FUNCTION_BLOCK FB_ScalingOffset_1
(*

The function block used to scaling input signal.

Constructor: 		Patryk Panylo
Company:		E. Riexinger GmbH
Date:			04.08.2015
Version:			1.00

Date:			Revision:		Who:				Comment
dd.mm.yyyy		x.xx			Initials			comment

*)
VAR_INPUT
	(* Input variables / Eingang Variablen *)
	bEnable							:BOOL;						(* Function block enable *)
	lrInput							:LREAL;						(* Input scaling proces value *)
	lrXLowLimit						:LREAL;						(* Upper limit of X range *)
	lrXUpperLimit						:LREAL; 						(*Upper limit of X range  *)
	lrYLowLimit						:LREAL; 						(* Low limit of Y range  *)
	lrYUpperLimit						:LREAL; 						(* Upper limit of Y range  *)
	usiPrecision						:USINT := 2; 					(* The number of digits after the decimal point depends on the requested precision *)
	lrOffset							:LREAL;						(* Offset of output *)
END_VAR
VAR_OUTPUT
	(* Output variables / Ausgang Variablen *)
	lrOutputRV						:LREAL;						(* Raw Value *)
	lrOutputPV						:LREAL;						(* Judgment Value  *)
END_VAR
VAR
	(* Instances / Instanzen *)
	fbScaling						:FB_Scaling;

	(* Enumerator  *)

	(* General flags / Allgemeine Variablen *)

END_VAR
VAR CONSTANT

END_VAR

IF NOT bEnable THEN
	fbScaling(
		bEnable := FALSE,
	);

	lrOutputRV := 0.0;					(* Raw Value *)
	lrOutputPV := 0.0;					(* Judgment Value *)
	RETURN;
END_IF

(* Scaling *)

fbScaling(
	bEnable := TRUE,
	lrInput := lrInput,
	lrXLowLimit := lrXLowLimit,
	lrXUpperLimit := lrXUpperLimit,
	lrYLowLimit := lrYLowLimit,
	lrYUpperLimit := lrYUpperLimit,
	usiPrecision := usiPrecision
);

lrOutputRV := fbScaling.lrOutputRV + lrOffset;
lrOutputPV := fbScaling.lrOutputPV + lrOffset;

END_FUNCTION_BLOCK

(* stored: Version 1.1.0.1, ProductVersion 3.1.4024.15
   POU FB_ScalingOffset_1: Id {5e2ee5e9-86f8-480b-bd1c-3ee2837effe7}, SpecialFunc None *)
